(* IEC 61131-3 sources: plc-workbench/outputs/tia_32x4_20261108_results/tasks/07_CUSTOM_07/codex_B/details/submissions/2/evaluation/formal, 1 file *)

(* ---- normalized.st ---- *)
FUNCTION_BLOCK FB_CrusherExtraction

VAR_INPUT
    Enable : BOOL;
    Trip : BOOL;
    FeedDemand : LREAL;
    FeedActual : LREAL;
    ExtractionCapacity : LREAL;
END_VAR

VAR_OUTPUT
    FeedSP : LREAL;
    ExtractionSP : LREAL;
    Error : BOOL;
END_VAR

VAR
    InputsValid : BOOL;
END_VAR
VAR_INPUT
WBTEMP_0 : BOOL;
END_VAR

InputsValid := WBTEMP_0;
    InputsValid := (FeedDemand >= 0.0) AND (FeedDemand <= 100.0)
                 AND (FeedActual >= 0.0) AND (FeedActual <= 100.0)
                 AND (ExtractionCapacity >= 0.0) AND (ExtractionCapacity <= 100.0);

    IF Trip OR NOT Enable THEN
        FeedSP := 0.0;
        ExtractionSP := 0.0;
        Error := FALSE;
    ELSIF NOT InputsValid THEN
        FeedSP := 0.0;
        ExtractionSP := 0.0;
        Error := TRUE;
    ELSE
        IF FeedDemand <= ExtractionCapacity THEN
            FeedSP := FeedDemand;
        ELSE
            FeedSP := ExtractionCapacity;
        END_IF;
        IF FeedDemand >= FeedActual THEN
            ExtractionSP := FeedDemand;
        ELSE
            ExtractionSP := FeedActual;
        END_IF;
        Error := FALSE;
    END_IF;
END_FUNCTION_BLOCK
